// TwinCAT 3 PLC project PLCStudent
// ProgramVersion: 3.1.4026.20
// libraries:
//   Tc2_Standard, * (Beckhoff Automation GmbH)
//   Tc2_System, * (Beckhoff Automation GmbH)
//   Tc3_Module, * (Beckhoff Automation GmbH)
// project tree:
//   / PlcTask.TcTTO
//   POUs/ ControlFBD.TcPOU, MAIN.TcPOU
// (motion and I/O tree: see PLC project plcsim)
// real-time tasks:
//   TASK PlcTask: cycle T#10ms, priority 20, ADS port 350
// variable links:
//   PLCSim/PLCSim Instance <-> PLCStudent/PLCStudent Instance
//     PlcTask Inputs/GVL.ixLed{1..8} <-> PlcTask Outputs/ControlFBD.qxLed{1..8}  (8 links)
//     PlcTask Outputs/GVL.qxButton{1..8} <-> PlcTask Inputs/ControlFBD.ixButton{1..8}  (8 links)

CONFIGURATION PLCStudent
    RESOURCE PLC ON TwinCAT3
        TASK PlcTask(INTERVAL := T#10ms, PRIORITY := 20);
        PROGRAM MAIN WITH PlcTask : MAIN;
    END_RESOURCE
END_CONFIGURATION

// ---- POUs/MAIN.TcPOU
PROGRAM MAIN
VAR
END_VAR

ControlFBD();

END_PROGRAM

// ---- POUs/ControlFBD.TcPOU
PROGRAM ControlFBD
VAR
	
	ixButton1 AT %I* : BOOL;
	ixButton2 AT %I* : BOOL;
	ixButton3 AT %I* : BOOL;
	ixButton4 AT %I* : BOOL;
	ixButton5 AT %I* : BOOL;
	ixButton6 AT %I* : BOOL;
	ixButton7 AT %I* : BOOL;
	ixButton8 AT %I* : BOOL;
	
	mxTime1:BOOL;
	mxTime2:BOOL;
	mxTime3:BOOL;
	mxTime4:BOOL;
	mxTime5:BOOL;
	mxTime6:BOOL;
	mxTime7:BOOL;
	mxTime8:BOOL;
	mxTime9:BOOL;
	
	mxStart:BOOL;
	
	
	
	qxLed1 AT %Q* : BOOL;
	qxLed2 AT %Q* : BOOL;
	qxLed3 AT %Q* : BOOL;
	qxLed4 AT %Q* : BOOL;
	qxLed5 AT %Q* : BOOL;
	qxLed6 AT %Q* : BOOL;
	qxLed7 AT %Q* : BOOL;
	qxLed8 AT %Q* : BOOL;

	fbTime1: TON;
	fbTime2: TON;
	fbTime3: TON;
	fbTime4: TON;
	fbTime5: TON;
	fbTime6: TON;
	fbTime7: TON;
	fbTime8: TON;
	fbTime9: TON;
	mxReturn: BOOL;
END_VAR
VAR // added by the converter: edge detectors and wires of the graphical bodies
    _w1, _w2, _w3, _w4, _w5, _w6, _w7 : BOOL;
END_VAR

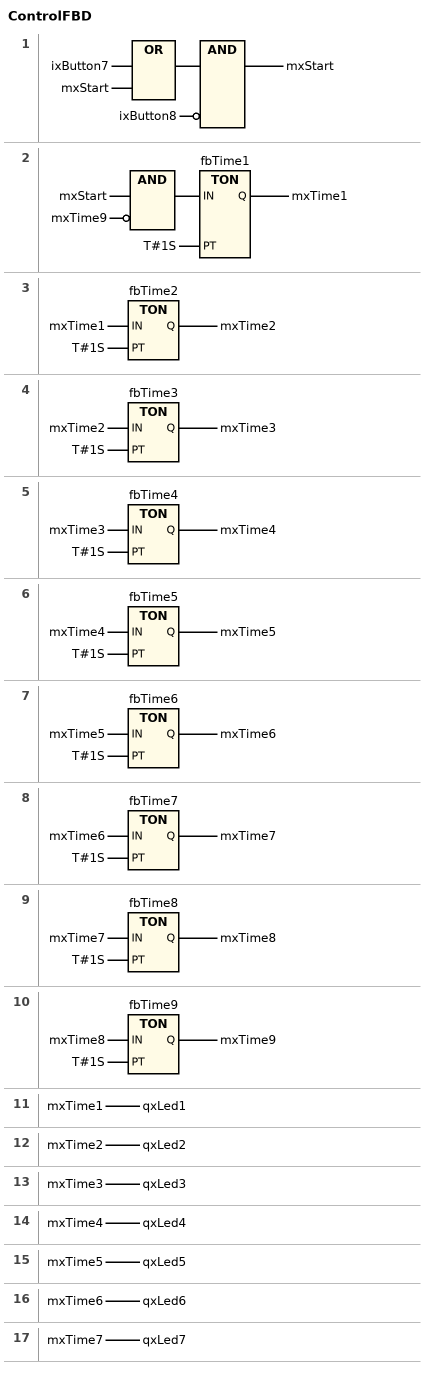
// NETWORK 1
mxStart := (ixButton7 OR mxStart) AND NOT ixButton8;

// NETWORK 2
fbTime1(IN := mxStart AND NOT mxTime9, PT := T#1S); // TON
mxTime1 := fbTime1.Q;

// NETWORK 3
fbTime2(IN := mxTime1, PT := T#1S); // TON
mxTime2 := fbTime2.Q;

// NETWORK 4
fbTime3(IN := mxTime2, PT := T#1S); // TON
mxTime3 := fbTime3.Q;

// NETWORK 5
fbTime4(IN := mxTime3, PT := T#1S); // TON
mxTime4 := fbTime4.Q;

// NETWORK 6
fbTime5(IN := mxTime4, PT := T#1S); // TON
mxTime5 := fbTime5.Q;

// NETWORK 7
fbTime6(IN := mxTime5, PT := T#1S); // TON
mxTime6 := fbTime6.Q;

// NETWORK 8
fbTime7(IN := mxTime6, PT := T#1S); // TON
mxTime7 := fbTime7.Q;

// NETWORK 9
fbTime8(IN := mxTime7, PT := T#1S); // TON
mxTime8 := fbTime8.Q;

// NETWORK 10
fbTime9(IN := mxTime8, PT := T#1S); // TON
mxTime9 := fbTime9.Q;

// NETWORK 11
qxLed1 := mxTime1;

// NETWORK 12
qxLed2 := mxTime2;

// NETWORK 13
qxLed3 := mxTime3;

// NETWORK 14
qxLed4 := mxTime4;

// NETWORK 15
qxLed5 := mxTime5;

// NETWORK 16
qxLed6 := mxTime6;

// NETWORK 17
qxLed7 := mxTime7;

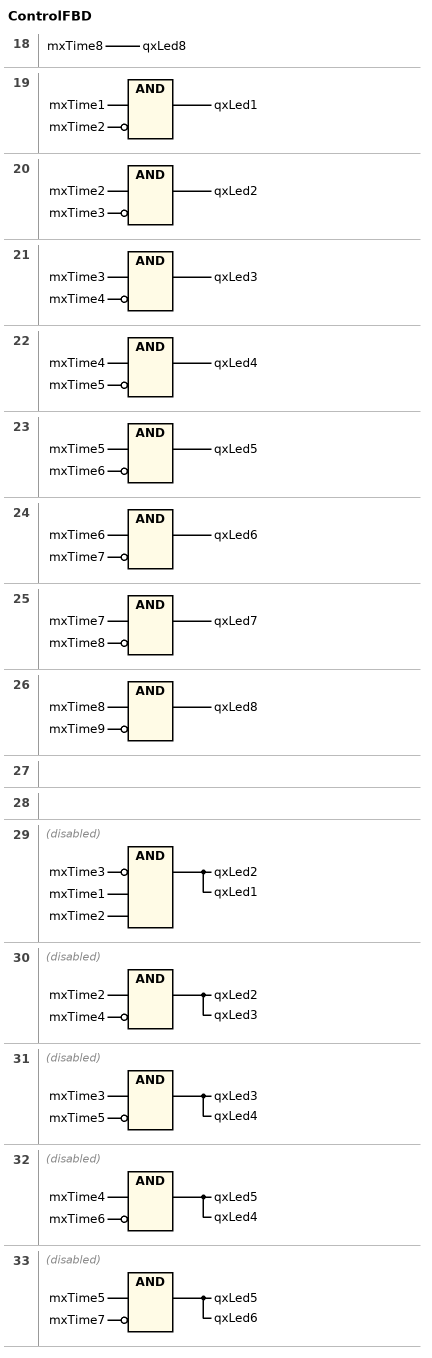
// NETWORK 18
qxLed8 := mxTime8;

// NETWORK 19
qxLed1 := mxTime1 AND NOT mxTime2;

// NETWORK 20
qxLed2 := mxTime2 AND NOT mxTime3;

// NETWORK 21
qxLed3 := mxTime3 AND NOT mxTime4;

// NETWORK 22
qxLed4 := mxTime4 AND NOT mxTime5;

// NETWORK 23
qxLed5 := mxTime5 AND NOT mxTime6;

// NETWORK 24
qxLed6 := mxTime6 AND NOT mxTime7;

// NETWORK 25
qxLed7 := mxTime7 AND NOT mxTime8;

// NETWORK 26
qxLed8 := mxTime8 AND NOT mxTime9;

// NETWORK 27

// NETWORK 28

// NETWORK 29 (disabled)
// _w1 := NOT mxTime3 AND mxTime1 AND mxTime2;
// qxLed2 := _w1;
// qxLed1 := _w1;

// NETWORK 30 (disabled)
// _w2 := mxTime2 AND NOT mxTime4;
// qxLed2 := _w2;
// qxLed3 := _w2;

// NETWORK 31 (disabled)
// _w3 := mxTime3 AND NOT mxTime5;
// qxLed3 := _w3;
// qxLed4 := _w3;

// NETWORK 32 (disabled)
// _w4 := mxTime4 AND NOT mxTime6;
// qxLed5 := _w4;
// qxLed4 := _w4;

// NETWORK 33 (disabled)
// _w5 := mxTime5 AND NOT mxTime7;
// qxLed5 := _w5;
// qxLed6 := _w5;

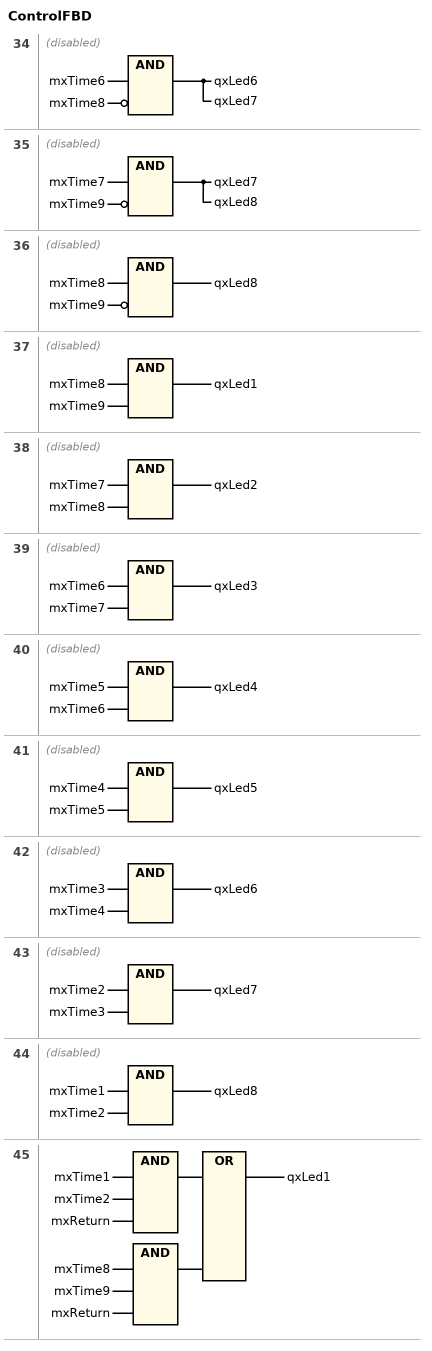
// NETWORK 34 (disabled)
// _w6 := mxTime6 AND NOT mxTime8;
// qxLed6 := _w6;
// qxLed7 := _w6;

// NETWORK 35 (disabled)
// _w7 := mxTime7 AND NOT mxTime9;
// qxLed7 := _w7;
// qxLed8 := _w7;

// NETWORK 36 (disabled)
// qxLed8 := mxTime8 AND NOT mxTime9;

// NETWORK 37 (disabled)
// qxLed1 := mxTime8 AND mxTime9;

// NETWORK 38 (disabled)
// qxLed2 := mxTime7 AND mxTime8;

// NETWORK 39 (disabled)
// qxLed3 := mxTime6 AND mxTime7;

// NETWORK 40 (disabled)
// qxLed4 := mxTime5 AND mxTime6;

// NETWORK 41 (disabled)
// qxLed5 := mxTime4 AND mxTime5;

// NETWORK 42 (disabled)
// qxLed6 := mxTime3 AND mxTime4;

// NETWORK 43 (disabled)
// qxLed7 := mxTime2 AND mxTime3;

// NETWORK 44 (disabled)
// qxLed8 := mxTime1 AND mxTime2;

// NETWORK 45
qxLed1 := mxTime1 AND mxTime2 AND mxReturn OR mxTime8 AND mxTime9 AND mxReturn;

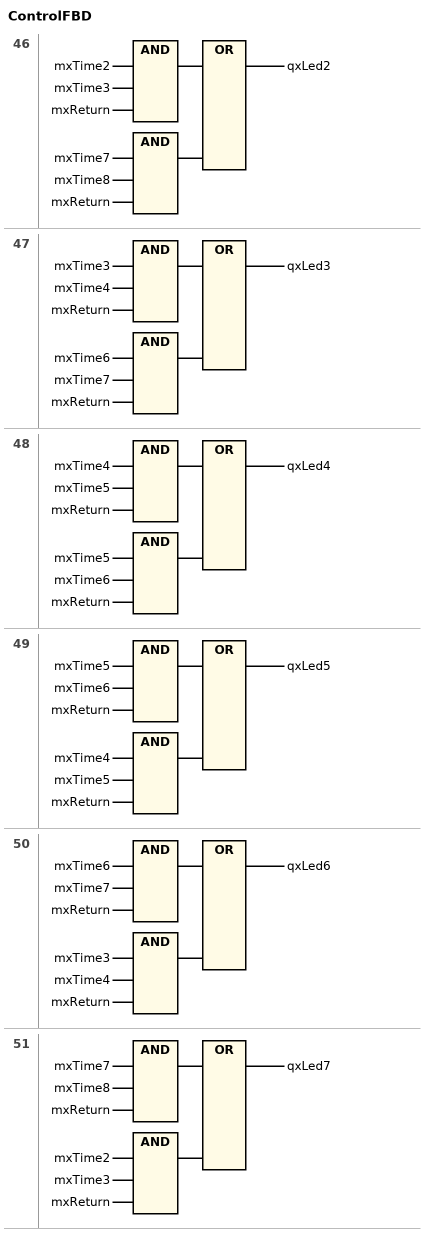
// NETWORK 46
qxLed2 := mxTime2 AND mxTime3 AND mxReturn OR mxTime7 AND mxTime8 AND mxReturn;

// NETWORK 47
qxLed3 := mxTime3 AND mxTime4 AND mxReturn OR mxTime6 AND mxTime7 AND mxReturn;

// NETWORK 48
qxLed4 := mxTime4 AND mxTime5 AND mxReturn OR mxTime5 AND mxTime6 AND mxReturn;

// NETWORK 49
qxLed5 := mxTime5 AND mxTime6 AND mxReturn OR mxTime4 AND mxTime5 AND mxReturn;

// NETWORK 50
qxLed6 := mxTime6 AND mxTime7 AND mxReturn OR mxTime3 AND mxTime4 AND mxReturn;

// NETWORK 51
qxLed7 := mxTime7 AND mxTime8 AND mxReturn OR mxTime2 AND mxTime3 AND mxReturn;

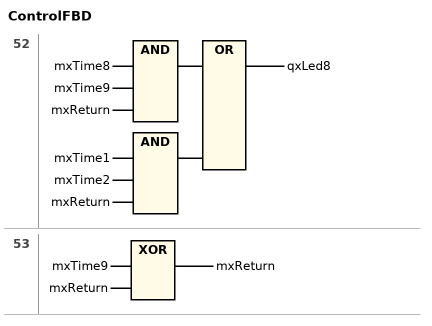
// NETWORK 52
qxLed8 := mxTime8 AND mxTime9 AND mxReturn OR mxTime1 AND mxTime2 AND mxReturn;

// NETWORK 53
mxReturn := mxTime9 XOR mxReturn;

END_PROGRAM
